Staubli VAL3: setReferencePos.pgx

public program setReferencePos(jointRx x_jPoint, num x_nDeviate)
// // 定义一个参考位置
// // x_jPoint: 设定的参考位置的值
// // x_nDeviate: 相对于reference point，允许的误差
begin
  // ---------------------------------------------------------------------------- //
  // 定义一个参考位置
  // x_jPoint: 设定的参考位置的值
  // x_nDeviate: 相对于reference point，允许的误差
  // ---------------------------------------------------------------------------- //
  jRefPoint=x_jPoint
  nRefDeviate=x_nDeviate
end
